FUNCTION_BLOCK SKILL_Gate (* The front desk of a skill, inside SKILL_Core: answers a client's Start, Stop, Abort or Reset at once (only the module's owner; Start only with the module in Execute, the skill not running, the values in range and the equipment free) and passes an accepted command on to SKILL_Control, as a parent's command is passed on. Technical: Decides a client's Start/Stop/Abort/Reset (owner only; Start only in module Execute, not running, parameters in range, equipment free) and passes accepted ones and a parent's on as GO_START, GO_HALT, GO_ABORT, GO_RESET to SKILL_Control *)
  (* Standard: 61499-2 *)
  (* Version 0.1, 2026-09-28, Project contributors, AAU Smart Production Lab *)
  PACKAGE modlib;
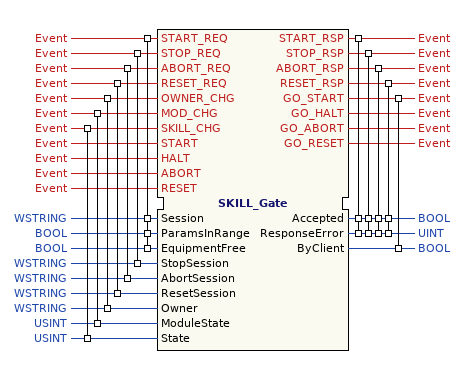
  EVENT_INPUT
    START_REQ WITH Session, ParamsInRange, EquipmentFree; (* Start(Session, parameters) was called: check Session, ParamsInRange, EquipmentFree *)
    STOP_REQ WITH StopSession; (* Stop(Session) was called *)
    ABORT_REQ WITH AbortSession; (* Abort(Session) was called *)
    RESET_REQ WITH ResetSession; (* Reset(Session) was called *)
    OWNER_CHG WITH Owner; (* The module's owner changed *)
    MOD_CHG WITH ModuleState; (* The module's state changed (its Stopping halts, its Aborting aborts the skill) *)
    SKILL_CHG WITH State; (* The skill's state changed (State, as SKILL_Control publishes it) *)
    START; (* The parent starts a run: passed on unchecked *)
    HALT; (* The parent stops the run: passed on unchecked *)
    ABORT; (* The parent aborts: passed on unchecked *)
    RESET; (* The parent resets: passed on unchecked *)
  END_EVENT
  EVENT_OUTPUT
    START_RSP WITH Accepted, ResponseError; (* Answer to Start *)
    STOP_RSP WITH Accepted, ResponseError; (* Answer to Stop *)
    ABORT_RSP WITH Accepted, ResponseError; (* Answer to Abort *)
    RESET_RSP WITH Accepted, ResponseError; (* Answer to Reset *)
    GO_START WITH ByClient; (* Start the run: a client's Start that was accepted, or the parent's (ByClient says which) *)
    GO_HALT; (* Stop the run: a client's Stop that was accepted, or the parent's HALT *)
    GO_ABORT; (* Abort: a client's Abort that was accepted, or the parent's ABORT *)
    GO_RESET; (* Reset: a client's Reset that was accepted, or the parent's RESET *)
  END_EVENT
  VAR_INPUT
    Session : WSTRING; (* Session ID of the caller of Start (must be the module's owner) *)
    ParamsInRange : BOOL; (* Every Start argument lies within its limits *)
    EquipmentFree : BOOL; (* The equipment is free, or held by this skill *)
    StopSession : WSTRING; (* Session ID of the caller of Stop *)
    AbortSession : WSTRING; (* Session ID of the caller of Abort *)
    ResetSession : WSTRING; (* Session ID of the caller of Reset *)
    Owner : WSTRING; (* Session ID of the module's owner (empty: free) *)
    ModuleState : USINT; (* PackML state: 1 Clearing, 2 Stopped, 3 Starting, 4 Idle, 6 Execute, 7 Stopping, 8 Aborting, 9 Aborted, 15 Resetting *)
    State : USINT; (* Skill state: 0 Idle, 1 Running, 2 Stopping, 3 Succeeded, 4 Failed, 5 Aborted *)
  END_VAR
  VAR_OUTPUT
    Accepted : BOOL; (* The call was accepted *)
    ResponseError : UINT; (* Why a call was refused (error code) *)
    ByClient : BOOL; (* The start came from a client over OPC UA (TRUE), or from the parent (FALSE) *)
  END_VAR
  VAR
    Owned : BOOL;
  END_VAR
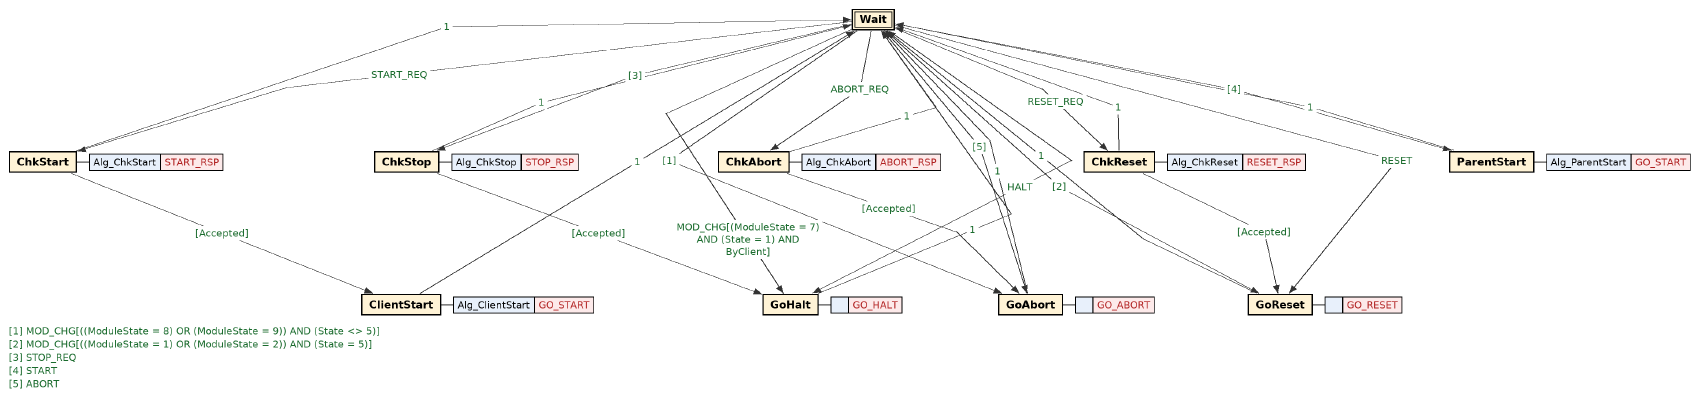
  EC_STATES
    Wait;
    ChkStart : Alg_ChkStart -> START_RSP;
    ChkStop : Alg_ChkStop -> STOP_RSP;
    ChkAbort : Alg_ChkAbort -> ABORT_RSP;
    ChkReset : Alg_ChkReset -> RESET_RSP;
    ClientStart : Alg_ClientStart -> GO_START;
    ParentStart : Alg_ParentStart -> GO_START;
    GoHalt : -> GO_HALT;
    GoAbort : -> GO_ABORT;
    GoReset : -> GO_RESET;
  END_STATES
  EC_TRANSITIONS
    Wait TO ChkStart := START_REQ;
    Wait TO ChkStop := STOP_REQ;
    Wait TO ChkAbort := ABORT_REQ;
    Wait TO ChkReset := RESET_REQ;
    Wait TO ParentStart := START;
    Wait TO GoHalt := HALT;
    Wait TO GoAbort := ABORT;
    Wait TO GoReset := RESET;
    Wait TO GoAbort := MOD_CHG[((ModuleState = 8) OR (ModuleState = 9)) AND (State <> 5)];
    Wait TO GoHalt := MOD_CHG[(ModuleState = 7) AND (State = 1) AND ByClient];
    Wait TO GoReset := MOD_CHG[((ModuleState = 1) OR (ModuleState = 2)) AND (State = 5)];
    ChkStart TO ClientStart := [Accepted];
    ChkStart TO Wait := 1;
    ChkStop TO GoHalt := [Accepted];
    ChkStop TO Wait := 1;
    ChkAbort TO GoAbort := [Accepted];
    ChkAbort TO Wait := 1;
    ChkReset TO GoReset := [Accepted];
    ChkReset TO Wait := 1;
    ClientStart TO Wait := 1;
    ParentStart TO Wait := 1;
    GoHalt TO Wait := 1;
    GoAbort TO Wait := 1;
    GoReset TO Wait := 1;
  END_TRANSITIONS
  ALGORITHM Alg_ChkStart IN ST:
Owned := (Session = Owner) AND (Owner <> "");
Accepted := FALSE;
IF NOT Owned THEN
  ResponseError := 5;
ELSIF ModuleState <> 6 THEN
  ResponseError := 4;
ELSIF (State = 1) OR (State = 2) THEN
  ResponseError := 6;
ELSIF State = 5 THEN
  ResponseError := 4;
ELSIF NOT ParamsInRange THEN
  ResponseError := 8;
ELSIF NOT EquipmentFree THEN
  ResponseError := 6;
ELSE
  Accepted := TRUE;
  ResponseError := 0;
END_IF;
  END_ALGORITHM
  ALGORITHM Alg_ChkStop IN ST:
Owned := (StopSession = Owner) AND (Owner <> "");
Accepted := Owned AND (State = 1);
IF NOT Owned THEN
  ResponseError := 5;
ELSIF NOT Accepted THEN
  ResponseError := 4;
ELSE
  ResponseError := 0;
END_IF;
  END_ALGORITHM
  ALGORITHM Alg_ChkAbort IN ST:
Owned := (AbortSession = Owner) AND (Owner <> "");
Accepted := Owned AND (State <> 5);
IF NOT Owned THEN
  ResponseError := 5;
ELSIF NOT Accepted THEN
  ResponseError := 4;
ELSE
  ResponseError := 0;
END_IF;
  END_ALGORITHM
  ALGORITHM Alg_ChkReset IN ST:
Owned := (ResetSession = Owner) AND (Owner <> "");
Accepted := Owned AND (State = 5);
IF NOT Owned THEN
  ResponseError := 5;
ELSIF NOT Accepted THEN
  ResponseError := 4;
ELSE
  ResponseError := 0;
END_IF;
  END_ALGORITHM
  ALGORITHM Alg_ClientStart IN ST:
ByClient := TRUE;
  END_ALGORITHM
  ALGORITHM Alg_ParentStart IN ST:
ByClient := FALSE;
  END_ALGORITHM
END_FUNCTION_BLOCK
